// TIA Portal V21 export
Screen "FP_Source"  NonexNone, Number=599
  ScreenLayer "Layer_0"
    Rectangle "FP_Frame" at 10,10 size 300x150
    Rectangle "FP_Status" at 20,20 size 60x40
      RangeAppearanceAnimation "RangeAppearanceAnimation"
        tag D_Range
        0..9: back #ff0000, fore #ffffff
        10..49: back #00a000, fore #000000
        50..99: back #0000ff, fore #ffff00
    IOField "FP_Value" at 100,20 size 100x30  FormatPattern=s99999
      ProcessValue := D_Int
    Bar "FP_Bar" at 220,20 size 30x130
      ProcessValue := D_Pct
    Circle "FP_Lamp" at 260,20 size 40x40
      SingleBitVisibilityAnimation "VisibilityAnimation"
        tag D_Vis
    TextField "FP_Title" at 20,120 size 180x20  Text="<body><p>Faceplate FP_C05</p></body>"
